{region 'Documentation'}
(*!
<summary>Check that the token count equals Expected.</summary>
<description>

StartIndex is an absolute declared IN index, not an offset. Length selects 1..255
elements; the complete selected range must fit IN. Invalid references or ranges report
Error.

Keep supplied arrays stable for the call. Input data is read, not copied or retained as a
snapshot.

Counts the currently selected region on evaluation, not occurrences across cycles.
TokenCount exposes the last computed count.

Token is the complete nonempty array pattern starting at its own lower bound and must fit
the selected search range; otherwise Error. Array token matching is exact.

Matches do not overlap: searching resumes after the whole matched token.

</description>
*)
{endregion}
FUNCTION_BLOCK AssertArrayTokenCntEqual_Byte EXTENDS AssertionBase
VAR_INPUT
    StartIndex : DINT; //! First selected index in IN; uses the array's declared index range, not a zero-based offset.
    Length : USINT; //! Number of selected elements starting at StartIndex; must fit the array range; valid range 1..255.
    Expected : UINT; //! Reference count for the named relation; counts occurrences, not array indices.
END_VAR
VAR_IN_OUT CONSTANT
    IN : ARRAY[*] OF BYTE; //! Keep the searched data stable during the call.
    Token : ARRAY[*] OF BYTE; //! Read-only nonempty token; keep stable during the call and within the selected search length.
END_VAR
VAR
    FTokenCount : UINT;
END_VAR

SUPER^();

{region 'Documentation'}
(*!
<summary>Validate configuration, count tokens and apply the count predicate.</summary>
*)
{endregion}
METHOD PROTECTED Assert
VAR
    InLowerIndex : DINT;
    InUpperIndex : DINT;
    EndIndex : LINT;
    TokenLowerIndex : DINT;
    TokenUpperIndex : DINT;
    TokenLength : LINT;
    Message : STRING(GVL_Constants.MessageLength);
END_VAR
IF NOT EvaluationActive THEN
    RETURN;
END_IF;

IF Result = E_Result.Error THEN
    RETURN;
END_IF;

// C0371: FB input is checked before any reference access.
{warning disable C0371}
IF NOT __ISVALIDREF(IN) THEN
    FTokenCount := 0;
    Error(Message := 'Assertion error: IN reference is invalid.');
    RETURN;
END_IF;

IF NOT __ISVALIDREF(Token) THEN
    FTokenCount := 0;
    Error(Message := 'Assertion error: Token reference is invalid.');
    RETURN;
END_IF;

TokenLowerIndex := LOWER_BOUND(Token, 1);
TokenUpperIndex := UPPER_BOUND(Token, 1);
TokenLength := DINT_TO_LINT(TokenUpperIndex) - DINT_TO_LINT(TokenLowerIndex) + 1;
IF (TokenLength <= 0) OR (TokenLength > USINT_TO_LINT(Length)) THEN
    FTokenCount := 0;
    Message := CONCAT('Assertion error: invalid token length. TokenLength = ',
        LINT_TO_STRING(TokenLength));
    Message := CONCAT(Message, ', Length = ');
    Message := CONCAT(Message, USINT_TO_STRING(Length));
    Error(Message := Message);
    RETURN;
END_IF;

InLowerIndex := LOWER_BOUND(IN, 1);
InUpperIndex := UPPER_BOUND(IN, 1);
EndIndex := DINT_TO_LINT(StartIndex) + USINT_TO_LINT(Length) - 1;
IF (Length = 0)
    OR (StartIndex < InLowerIndex) OR (StartIndex > InUpperIndex)
    OR (EndIndex > DINT_TO_LINT(InUpperIndex)) THEN
    FTokenCount := 0;
    Message := CONCAT('Assertion error: invalid search range. StartIndex = ',
        DINT_TO_STRING(StartIndex));
    Message := CONCAT(Message, ', Length = ');
    Message := CONCAT(Message, USINT_TO_STRING(Length));
    Error(Message := Message);
    RETURN;
END_IF;

IF Result = E_Result.Failed THEN
    RETURN;
END_IF;

FTokenCount := CountArrayTokens_Byte(StartIndex := StartIndex,
    Length := Length,
    Token := Token,
    IN := IN);

IF FTokenCount <> Expected THEN
    Message := CONCAT('Assertion failed: array token count violates Equal. Actual = ',
        UINT_TO_STRING(FTokenCount));
    Message := CONCAT(Message, ', Expected = ');
    Message := CONCAT(Message, UINT_TO_STRING(Expected));
    Message := CONCAT(Message, ', TokenRange = [');
    Message := CONCAT(Message, DINT_TO_STRING(TokenLowerIndex));
    Message := CONCAT(Message, '..');
    Message := CONCAT(Message, DINT_TO_STRING(TokenUpperIndex));
    Message := CONCAT(Message, ']');
    Fail(Message := Message);
    RETURN;
END_IF;

Pass();
{warning restore C0371}
END_METHOD

{region 'Documentation'}
(*!
<summary>Clear the retained count on framework reset.</summary>
*)
{endregion}
METHOD PROTECTED ResetAssertion
FTokenCount := 0;
END_METHOD

{region 'Documentation'}
(*!
<summary>Return the most recently evaluated token count.</summary>
<description>

Counts occurrences in one selected array region, not across PLC cycles. Retained while
disabled or after Failed; reset and detected configuration errors clear it. Reading this
property does not search the array.

</description>
*)
{endregion}
{attribute 'monitoring' := 'call'}
PROPERTY PUBLIC TokenCount : UINT //! Return the most recently evaluated token count.
GET // PUBLIC
TokenCount := FTokenCount;
END_GET
END_PROPERTY

END_FUNCTION_BLOCK

(* stored: Version 1.1.0.1
   POU AssertArrayTokenCntEqual_Byte: Id {b151da34-1c73-4ec6-bd9b-b0cd8b9864f7}, SpecialFunc None
   Folder Internal: Id {c6c8a7f7-5df8-43e3-b064-b91c309645cb}
   Method Assert: Id {2ba0bd2f-b17f-4c24-9cfa-8d097c6c50b6}
   Method ResetAssertion: Id {337af9e2-ba5d-46a3-ab97-770713429371}
   Property TokenCount: Id {60048750-cec6-496d-a3cc-90b99848ddc5}
   Get Get: Id {4f21430b-1a8e-4262-b841-e73f74ed22be} *)
